// TIA Portal project "S71200_v1" (V16)

(* hardware
DEVICE "S7-1200 station_1"  S7-1200 Station
   slot 0: "Rack_0"  S7-1200 Rack  Rack  V1.0
   slot 1: "PLC_1"  CPU 1212C AC/DC/Rly  6ES7 212-1BE40-0XB0  V4.4
DEVICE "GSD device_2"  GSD.Device.PN
   slot 0: "Rack"  Rack  V1.0
   slot 0: "BannerSafetyController"  Banner Safety Controller  Banner-Safety-Controller
      slot 0: "Submodule 1"  Submodule 1
      slot 1: "I"  I
         slot 1: "P1"  P1
      slot 1: "4 Status Bytes, Bits 0..31_1"  4 Status Bytes, Bits 0..31  1.0
         slot 0: "4 Status Bytes, Bits 0..31"  4 Status Bytes, Bits 0..31
      slot 2: "4 Status Bytes, Bits 0..31_2"  4 Status Bytes, Bits 0..31  1.0
         slot 0: "4 Status Bytes, Bits 0..31"  4 Status Bytes, Bits 0..31
      slot 3: "4 Status Bytes, Bits 0..31_3"  4 Status Bytes, Bits 0..31  1.0
         slot 0: "4 Status Bytes, Bits 0..31"  4 Status Bytes, Bits 0..31
      slot 4: "4 Status Bytes, Bits 0..31_4"  4 Status Bytes, Bits 0..31  1.0
         slot 0: "4 Status Bytes, Bits 0..31"  4 Status Bytes, Bits 0..31
      slot 5: "4 Status Bytes, Bits 0..31_5"  4 Status Bytes, Bits 0..31  1.0
         slot 0: "4 Status Bytes, Bits 0..31"  4 Status Bytes, Bits 0..31
      slot 6: "4 Status Bytes, Bits 0..31_6"  4 Status Bytes, Bits 0..31  1.0
         slot 0: "4 Status Bytes, Bits 0..31"  4 Status Bytes, Bits 0..31
      slot 7: "4 Status Bytes, Bits 0..31_7"  4 Status Bytes, Bits 0..31  1.0
         slot 0: "4 Status Bytes, Bits 0..31"  4 Status Bytes, Bits 0..31
      slot 8: "4 Status Bytes, Bits 0..31_8"  4 Status Bytes, Bits 0..31  1.0
         slot 0: "4 Status Bytes, Bits 0..31"  4 Status Bytes, Bits 0..31
      slot 9: "4 Status Bytes, Bits 0..31_9"  4 Status Bytes, Bits 0..31  1.0
         slot 0: "4 Status Bytes, Bits 0..31"  4 Status Bytes, Bits 0..31
      slot 10: "4 Status Bytes, Bits 0..31_10"  4 Status Bytes, Bits 0..31  1.0
         slot 0: "4 Status Bytes, Bits 0..31"  4 Status Bytes, Bits 0..31
      slot 11: "4 Status Bytes, Bits 0..31_11"  4 Status Bytes, Bits 0..31  1.0
         slot 0: "4 Status Bytes, Bits 0..31"  4 Status Bytes, Bits 0..31
      slot 12: "4 Status Bytes, Bits 0..31_12"  4 Status Bytes, Bits 0..31  1.0
         slot 0: "4 Status Bytes, Bits 0..31"  4 Status Bytes, Bits 0..31
      slot 13: "8 Bytes Virtual On/Off/ME Data_1"  8 Bytes Virtual On/Off/ME Data  1.0
         slot 0: "Subslot 1 On/Off Data"  Subslot 1 On/Off Data
      slot 14: "2 Bytes RCD Data_1"  2 Bytes RCD Data  1.0
         slot 0: "Subslot 1 Reset/Cancel Delay Data"  Subslot 1 Reset/Cancel Delay Data
      slot 15: "2 Byte RCD Acutation Code_1"  2 Byte RCD Acutation Code  1.0
         slot 0: "Subslot 1 RCD Enable"  Subslot 1 RCD Enable
      slot 16: "RCD Data Feedback Register_1"  RCD Data Feedback Register  1.0
         slot 0: "Subslot 1 RCD Data Feedback"  Subslot 1 RCD Data Feedback
      slot 17: "RCD Passcode Feedback Register_1"  RCD Passcode Feedback Register  1.0
         slot 0: "Subslot 1 RCD Passcode Feedback"  Subslot 1 RCD Passcode Feedback
*)

// ===== PLC "PLC_1"  CPU 1212C AC/DC/Rly =====

VAR_GLOBAL   // PLC tag table "Default tag table"
   "Clock_Byte" AT %MB0 : Byte;
   "Clock_10Hz" AT %M0.0 : Bool;
   "Clock_5Hz" AT %M0.1 : Bool;
   "Clock_2.5Hz" AT %M0.2 : Bool;
   "Clock_2Hz" AT %M0.3 : Bool;
   "Clock_1.25Hz" AT %M0.4 : Bool;
   "Clock_1Hz" AT %M0.5 : Bool;
   "Clock_0.625Hz" AT %M0.6 : Bool;
   "Clock_0.5Hz" AT %M0.7 : Bool;
END_VAR

VAR_GLOBAL   // PLC tag table "Banner"
   "SC10_ManualResetRequired" AT %I1.0 : Bool;
   "SC10_RO1Status" AT %I37.0 : Bool;
   "SC10_RO2Status" AT %I37.1 : Bool;
   "PLC_VirtualNonSafetyOutput" AT %Q64.0 : Bool;
   "SC10_MagSwitchStatus" AT %I17.0 : Bool;
   "SC10_DoorSwitchStatus" AT %I17.1 : Bool;
   "SC10_EmStopStatus" AT %I17.2 : Bool;
   "PLC_BypassMagSwitch" AT %Q64.1 : Bool;
END_VAR

VAR_GLOBAL   // PLC tag table "FIO"
   "FIO_MCStart" AT %Q1.0 : Bool;
   "FIO_MCStop" AT %Q1.1 : Bool;
   "FIO_BypassMagSwitch" AT %I200.0 : Bool;
   "FIO_Em-Stop" AT %I200.1 : Bool;
END_VAR

FUNCTION "Banner" : Void   // FC1, SCL
{ S7_Optimized_Access := 'TRUE' }
VERSION : 0.1
   VAR_INPUT
      SC10_RO1Status : Bool;
      SC10_RO2Status : Bool;
      FIO_MuteMagSwitch : Bool;
      FIO_EmStop : Bool;
   END_VAR
   VAR_OUTPUT
      FIO_MCStart : Bool;
      FIO_MCStop : Bool;
      PLC_BypassMagSwitch : Bool;
      PLC_VirtualNonSafetyOutput : Bool;
   END_VAR
BEGIN
   //Using relay outptus to control Machine center
   IF #SC10_RO1Status AND #SC10_RO2Status THEN
       #FIO_MCStart := true;
       #FIO_MCStop := false;
   ELSE
       #FIO_MCStart := false;
       #FIO_MCStop := true;
   END_IF;

   //Muting Magnetic sensor
   #PLC_BypassMagSwitch := #FIO_MuteMagSwitch;

   //PLC E-Stop to Virtual non safety input of SC10
   #PLC_VirtualNonSafetyOutput := #FIO_EmStop;
END_FUNCTION

ORGANIZATION_BLOCK "Main"   // OB1, LAD, ProgramCycle
TITLE = "Main Program Sweep (Cycle)"
{ S7_Optimized_Access := 'TRUE' }
VERSION : 0.1
   VAR_INPUT
      Initial_Call : Bool;   // Initial call of this OB
      Remanence : Bool;   // =True, if remanent data are available
   END_VAR
BEGIN

REGION Network 1
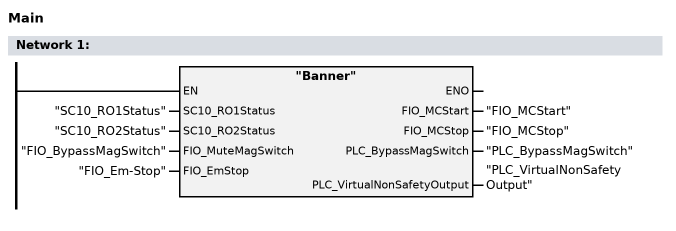
   RUNG wire#powerrail
      "Banner"(SC10_RO1Status := "SC10_RO1Status", SC10_RO2Status := "SC10_RO2Status", FIO_MuteMagSwitch := "FIO_BypassMagSwitch", FIO_EmStop := "FIO_Em-Stop", FIO_MCStart => "FIO_MCStart", FIO_MCStop => "FIO_MCStop", PLC_BypassMagSwitch => "PLC_BypassMagSwitch", PLC_VirtualNonSafetyOutput => "PLC_VirtualNonSafetyOutput")
   END_RUNG
   // the same network as SCL:
   "Banner"(SC10_RO1Status := "SC10_RO1Status",
            SC10_RO2Status := "SC10_RO2Status",
            FIO_MuteMagSwitch := "FIO_BypassMagSwitch",
            FIO_EmStop := "FIO_Em-Stop",
            FIO_MCStart => "FIO_MCStart",
            FIO_MCStop => "FIO_MCStop",
            PLC_BypassMagSwitch => "PLC_BypassMagSwitch",
            PLC_VirtualNonSafetyOutput => "PLC_VirtualNonSafetyOutput");
END_REGION
END_ORGANIZATION_BLOCK